{region 'Documentation'}
(*!
<summary>Checks Parallel registration order and shared slot across negative array bounds.</summary>
<description>Child mocks are inert interface identities and slot storage only; no child initialization or FB call is performed.</description>
*)
{endregion}
FUNCTION_BLOCK Test_SuiteBuilderParallel EXTENDS TestCaseBase
VAR
    FBuilder : TestSuiteConfigurationBuilder;
    FCases : ARRAY[-2..1] OF I_TestCase;
    FChildA : TestCaseMock;
    FChildB : TestCaseMock;
    FScenarioExecuted : BOOL;
    FChecksEvaluated : BOOL;
    FRegistration : AssertTrue;
    FRegistrationMatches : BOOL;
    FOrder : AssertTrue;
    FOrderMatches : BOOL;
    FSlots : AssertTrue;
    FSlotsMatches : BOOL;
    FMetadata : AssertTrue;
    FMetadataMatches : BOOL;
    FFinalization : AssertTrue;
    FFinalizationMatches : BOOL;
END_VAR

SUPER^();

{region 'Documentation'}
(*!
<summary>Contributes each owned Assertion once without executing it.</summary>
*)
{endregion}
METHOD PROTECTED AggregateResults
VAR_INPUT
    Aggregator : I_ResultAggregator; //! Borrowed result sink owned by the outer Test Case; add this test's checking Assertions without resetting or retaining the sink.
END_VAR
Aggregator.AddProvider(Provider := FRegistration);
Aggregator.AddProvider(Provider := FOrder);
Aggregator.AddProvider(Provider := FSlots);
Aggregator.AddProvider(Provider := FMetadata);
Aggregator.AddProvider(Provider := FFinalization);
END_METHOD

{region 'Documentation'}
(*!
<summary>Requires successful base and owned Assertion initialization.</summary>
*)
{endregion}
METHOD PROTECTED CheckInitialization : BOOL //! TRUE when the inherited initialization check and this concrete fixture check both accept the setup.
CheckInitialization := FALSE;
IF NOT SUPER^.CheckInitialization() THEN
    RETURN;
END_IF;

CheckInitialization := FRegistration.IsInitialized
    AND FOrder.IsInitialized
    AND FSlots.IsInitialized
    AND FMetadata.IsInitialized
    AND FFinalization.IsInitialized;
END_METHOD

{region 'Documentation'}
(*!
<summary>Configures one direct builder scenario and its named Assertions.</summary>
*)
{endregion}
METHOD PROTECTED Configure
FPreparationStateCount := 0;
FTestStateCount := 1;
FScenarioExecuted := FALSE;
FChecksEvaluated := FALSE;

FRegistrationMatches := FALSE;
FRegistration.Initialize(Parent := THIS^,
    AssertionName := 'Registration');
FOrderMatches := FALSE;
FOrder.Initialize(Parent := THIS^,
    AssertionName := 'Order');
FSlotsMatches := FALSE;
FSlots.Initialize(Parent := THIS^,
    AssertionName := 'Slots');
FMetadataMatches := FALSE;
FMetadata.Initialize(Parent := THIS^,
    AssertionName := 'Metadata');
FFinalizationMatches := FALSE;
FFinalization.Initialize(Parent := THIS^,
    AssertionName := 'Finalization');
END_METHOD

{region 'Documentation'}
(*!
<summary>Completes Abort immediately; no asynchronous resource operation is started.</summary>
*)
{endregion}
METHOD PROTECTED ProcessAbort
VAR_INPUT
    Enable : BOOL; //! Phase permission supplied by the owning Test Case; FALSE does not authorize progression, while observation may continue.
END_VAR
IF Enable THEN
    CompleteAbort();
END_IF;
END_METHOD

{region 'Documentation'}
(*!
<summary>Evaluates recorded observations and consumes pending resets on disabled calls.</summary>
*)
{endregion}
METHOD PROTECTED ProcessAssertions
VAR_INPUT
    Enable : BOOL; //! Phase permission supplied by the owning Test Case; FALSE does not authorize progression, while observation may continue.
END_VAR
FRegistration(Enable := Enable,
    State := State,
    IN := FRegistrationMatches);

FOrder(Enable := Enable,
    State := State,
    IN := FOrderMatches);

FSlots(Enable := Enable,
    State := State,
    IN := FSlotsMatches);

FMetadata(Enable := Enable,
    State := State,
    IN := FMetadataMatches);

FFinalization(Enable := Enable,
    State := State,
    IN := FFinalizationMatches);

IF Enable AND FRegistration.EvaluationActive
    AND FOrder.EvaluationActive
    AND FSlots.EvaluationActive
    AND FMetadata.EvaluationActive
    AND FFinalization.EvaluationActive THEN
    FChecksEvaluated := TRUE;
END_IF;
END_METHOD

{region 'Documentation'}
(*!
<summary>No Preparation phase is needed for synchronous builder calls.</summary>
*)
{endregion}
METHOD PROTECTED ProcessPreparations
VAR_INPUT
    // SA0033: Required override signature; this scenario has no Preparation work.
    {attribute 'analysis' := '-33'}
    Enable : BOOL; //! Phase permission supplied by the owning Test Case; FALSE does not authorize progression, while observation may continue.
END_VAR
END_METHOD

{region 'Documentation'}
(*!
<summary>Clears recorded checks and Assertion results; each scenario initializes its own builder.</summary>
*)
{endregion}
METHOD PROTECTED ProcessReset
FScenarioExecuted := FALSE;
FChecksEvaluated := FALSE;
FRegistrationMatches := FALSE;
FRegistration.Reset();
FOrderMatches := FALSE;
FOrder.Reset();
FSlotsMatches := FALSE;
FSlots.Reset();
FMetadataMatches := FALSE;
FMetadata.Reset();
FFinalizationMatches := FALSE;
FFinalization.Reset();
CompleteReset();
END_METHOD

{region 'Documentation'}
(*!
<summary>Runs setup operations once, then completes after their observations have been evaluated.</summary>
*)
{endregion}
METHOD PROTECTED ProcessTests
VAR_INPUT
    Enable : BOOL; //! Phase permission supplied by the owning Test Case; FALSE does not authorize progression, while observation may continue.
END_VAR
IF NOT Enable THEN
    RETURN;
END_IF;

IF FChecksEvaluated THEN
    CompleteTests();
ELSIF NOT FScenarioExecuted THEN
    RunScenario();
    FScenarioExecuted := TRUE;
END_IF;
END_METHOD

{region 'Documentation'}
(*!
<summary>Checks Parallel registration order and shared slot across negative array bounds.</summary>
*)
{endregion}
METHOD PRIVATE RunScenario
VAR
    ChildA : I_TestCase;
    ChildB : I_TestCase;
    AcceptedA : BOOL;
    AcceptedB : BOOL;
    Config : ST_TestCaseCollectionConfig;
END_VAR
ChildA := FChildA;
ChildB := FChildB;
FBuilder.Initialize(Mode := E_OrchestrationMode.Parallel,
    TestCases := FCases);
AcceptedA := FBuilder.Register(TestCase := ChildB);
AcceptedB := FBuilder.Register(TestCase := ChildA);
FRegistrationMatches := AcceptedA AND AcceptedB;
FOrderMatches := (FCases[-2] = ChildB) AND (FCases[-1] = ChildA)
    AND (FCases[0] = 0) AND (FCases[1] = 0);
FSlotsMatches := (FChildA.ExecutionSlot = 1) AND (FChildB.ExecutionSlot = 1);
FMetadataMatches := (FBuilder.FirstIndex = -2) AND (FBuilder.LastIndex = 1)
    AND (FBuilder.Count = 2) AND (FBuilder.Mode = E_OrchestrationMode.Parallel);

Config := FBuilder.Finalize();
FFinalizationMatches := Config.IsValid AND FBuilder.IsValid AND FBuilder.IsFinalized
    AND (Config.FirstIndex = -2) AND (Config.LastIndex = 1) AND (Config.Count = 2)
    AND (Config.Mode = E_OrchestrationMode.Parallel);
END_METHOD

END_FUNCTION_BLOCK

(* stored: Version 1.1.0.1
   POU Test_SuiteBuilderParallel: Id {a78fd5a7-14ff-407d-873a-bc98b9e585a0}, SpecialFunc None
   Folder Internal: Id {00560001-0056-4056-8056-000000000016}
   Method AggregateResults: Id {00560001-0056-4056-8056-000000000014}
   Method CheckInitialization: Id {00560001-0056-4056-8056-00000000000d}
   Method Configure: Id {00560001-0056-4056-8056-00000000000c}
   Method ProcessAbort: Id {00560001-0056-4056-8056-00000000000f}
   Method ProcessAssertions: Id {00560001-0056-4056-8056-000000000013}
   Method ProcessPreparations: Id {00560001-0056-4056-8056-00000000000e}
   Method ProcessReset: Id {00560001-0056-4056-8056-000000000010}
   Method ProcessTests: Id {00560001-0056-4056-8056-000000000011}
   Method RunScenario: Id {00560001-0056-4056-8056-000000000012} *)
